Fanuc KAREL source: kc00018.KL

-- PROVISIONAL review KL for V940-1; original PC SHA256 d8d957c9dec6e45f9b679b51c2ebaf765fae3dc62dc094cf673abcce648b0100
-- Incomplete behavior may be omitted. Consult companion uncertainty JSON. Do not deploy.
PROGRAM KC00018
%NOLOCKGROUP
BEGIN
  -- V9_ZERO_TABLE_METADATA_HINT layout=0002_ascii; no indexed target words; source/name/runtime held
  -- UNRESOLVED_PC offsets 5-63; opcodes 27,22,2A,22,2A,22,22,2A,22,22,22,22,31
  -- UNRESOLVED_PC offsets 68-72; opcodes 7F
END KC00018
